(* IEC 61131-3 sources: STEPROBOT/docs/manual_control_r6_3/plc/reference, 5 files *)

(* ---- GVL_ManualBridge.st ---- *)
{attribute 'qualified_only'}
VAR_GLOBAL PERSISTENT RETAIN
    // PC extension: no overlap with HR200..215, HR300..363 or FTP HR6000+.
    aCommand AT %MW220 : ARRAY[0..15] OF WORD;
    aStatus AT %MW400 : ARRAY[0..31] OF WORD;
END_VAR
VAR_GLOBAL
    // Local configuration. Assign ONE unused GDI slot to manual_service before setting TRUE.
    xInstalled : BOOL := FALSE;
    xServiceBindingConfirmed : BOOL := FALSE;
    uiServiceProgram : UINT := 10;
    // PRG_ManualBridge is the only writer. PRG_RobotBridge reads these requests.
    xActive : BOOL;
    xStartRequest : BOOL;
    xStopRequest : BOOL;
END_VAR

(* ---- GVL_ManualPosition.st ---- *)
{attribute 'qualified_only'}
VAR_GLOBAL PERSISTENT RETAIN
    // Read-only position feedback to the PC. No robot or local permit writes.
    // MW450 requires both attributes. The bridge rebuilds this block every scan.
    aStatus AT %MW450 : ARRAY[0..39] OF WORD;
END_VAR

(* ---- GVL_ParamProbe.st ---- *)
{attribute 'qualified_only'}
VAR_GLOBAL
    // Mapped to existing ParamProbe_Write FC16 offset4 length4. Single writer: PRG_ManualBridge.
    aParamTx : ARRAY[0..3] OF WORD;
END_VAR

(* ---- GVL_RobotBridge.st ---- *)
// REFERENCE ONLY. Keep the field project declarations and boot counter; do not import.
{attribute 'qualified_only'}
VAR_GLOBAL PERSISTENT RETAIN
    // PC <-> PLC. Inovance native Modbus TCP slave: MWn <-> HR offset n.
    // Commission by reading HR300=16#4D42 and HR301=2 before permitting motion.
    aHostCmd AT %MW200 : ARRAY[0..15] OF WORD;
    aHostStatus AT %MW300 : ARRAY[0..63] OF WORD;

END_VAR

VAR_GLOBAL
    // PLC master -> STEP slave: FC04 / offset 0 / 32 WORD.
    aRobotRx : ARRAY[0..31] OF WORD;
    // PLC master -> STEP slave: ONE FC16 / offset 0 / 2 WORDs.
    // Map BOTH aRobotTx[0] and aRobotTx[1], NOT wRobotTxControl alone.
    aRobotTx : ARRAY[0..1] OF WORD;
    wRobotTxControl : WORD; // first-word diagnostic alias, not a separate channel

    // Local commissioning/operation inputs. Do not map these into aHostCmd.
    xCommissioned : BOOL := FALSE;
    // Set locally ONLY after checking DI49..56 and the GDI program bindings.
    xGdiProgramMappingConfirmed : BOOL := FALSE;
    xRemotePermit : BOOL := FALSE;
    // Optional native master/channel fault. FALSE leaves DO42 watchdog in use.
    xNativeModbusError : BOOL := FALSE;

    // Published live diagnostics.
    xRobotLinkOK : BOOL;
    xRobotRunning : BOOL;
    xRobotPaused : BOOL;
    xRobotStopped : BOOL;
    xRobotEnabled : BOOL;
    xRobotAlarm : BOOL;
    xRobotEmergency : BOOL;
    xRobotExternalAuto : BOOL;
    xHostRegistered : BOOL;
    xHostAlive : BOOL;
    xBusy : BOOL;
    xStopInterlock : BOOL;
    xLoadOperatorConfirmed : BOOL;
END_VAR

(* ---- GVL_RobotBridgeRetain.st ---- *)
// REFERENCE ONLY. Keep the field project declarations and boot counter; do not import.
{attribute 'qualified_only'}
VAR_GLOBAL PERSISTENT RETAIN
    // Incremented on application initialization, not on every scan.
    // Also require a fresh registration; a cold reset can reset RETAIN memory.
    udiBootCounter : UDINT := 0;
END_VAR
